(* IEC 61131-3 sources: T4Exjobb/Sigma/Stations/MachineControl/MachineControl/Class/_TCPIP_SERVER (part 2) *)

        (*================================================================*)
        else // - INVALID COMMAND
        (*================================================================*)
          Retcode := TCP_SVR_ERR_SET_PARA_INVALID_CMD;

      end_case;
    else
      Retcode := TCP_SVR_ERR_INVALID_SOCKET;
    end_if;
  else
    Retcode := TCP_SVR_ERR_INVALID_SOCKET;
  end_if;

END_FUNCTION

FUNCTION VIRTUAL GLOBAL _TCPIP_SERVER::ReadMainParameter
	VAR_INPUT
		Cmd 	: DINT;
		SubCmd 	: DINT;
		pParaValue 	: ^DINT;
	END_VAR
	VAR_OUTPUT
		Retcode 	: DINT;
	END_VAR

  Retcode := TCP_SVR_NO_ERROR;

  if (usInit > 0) then
    case Cmd of
      (*================================================================*)
      TCPSVR_CMD_SETSOCKOPT:
      (*================================================================*)
        case SubCmd of
          (*==================================================*)
          TCPSVR_SOCKOPT_NAGLE:
          (*==================================================*)
            if (MainSockOpt.Nagle = false) then
              pParaValue^ := 0;
            else
              pParaValue^ := 1;
            end_if;
          (*==================================================*)
          TCPSVR_SOCKOPT_KEEPALIVE:
          (*==================================================*)
            if (MainSockOpt.KeepAlive = false) then
              pParaValue^ := 0;
            else
              pParaValue^ := 1;
            end_if;
          (*==================================================*)
          TCPSVR_SOCKOPT_DELAYEDACK:
          (*==================================================*)
            if (MainSockOpt.DelayedAck = false) then
              pParaValue^ := 0;
            else
              pParaValue^ := 1;
            end_if;
          (*==================================================*)
          TCPSVR_SOCKOPT_REUSEADDR:
          (*==================================================*)
            if (MainSockOpt.ReuseAddr = false) then
              pParaValue^ := 0;
            else
              pParaValue^ := 1;
            end_if;
          (*==================================================*)
          else // - INVALID SUB COMMAND
          (*==================================================*)
            Retcode := TCP_SVR_ERR_SET_PARA_INVALID_SUB_CMD;
        end_case;

      (*================================================================*)
      TCPSVR_CMD_TASKPRIO:
      (*================================================================*)
        case SubCmd of
          (*==================================================*)
          TCPSVR_SUB_CMD_TASKPRIO:
          (*==================================================*)
            pParaValue^ := AP_TaskPriority$DINT;
          (*==================================================*)
          else // - INVALID SUB COMMAND
          (*==================================================*)
            Retcode := TCP_SVR_ERR_SET_PARA_INVALID_SUB_CMD;
        end_case;

      (*================================================================*)
      TCPSVR_CMD_KEEPALIVEPARA: // - ASYNC TASK PRIORITY
      (*================================================================*)
        case SubCmd of
          (*==================================================*)
          TCPSVR_KEEPALIVE_KEEPIDLE:
          (*==================================================*)
            pParaValue^ := KeepAlivePara.keepIDLE;
          (*==================================================*)
          TCPSVR_KEEPALIVE_KEEPINTVL:
          (*==================================================*)
            pParaValue^ := KeepAlivePara.keepINTVL;
          (*==================================================*)
          TCPSVR_KEEPALIVE_KEEPCNT:
          (*==================================================*)
            pParaValue^ := KeepAlivePara.keepCNT;
          (*==================================================*)
          else // - INVALID SUB COMMAND
          (*==================================================*)
            Retcode := TCP_SVR_ERR_SET_PARA_INVALID_SUB_CMD;
        end_case;

      (*================================================================*)
      TCPSVR_CMD_CLOSESOCKETTYPE:
      (*================================================================*)
        case SubCmd of
          (*==================================================*)
          TCPSVR_CLOSESOCKETTYPE:
          (*==================================================*)
            pParaValue^$UDINT := CloseSocketType;
          (*==================================================*)
          else // - INVALID SUB COMMAND
          (*==================================================*)
            Retcode := TCP_SVR_ERR_SET_PARA_INVALID_SUB_CMD;
        end_case;

      (*================================================================*)
      else // - INVALID COMMAND
      (*================================================================*)
        Retcode := TCP_SVR_ERR_SET_PARA_INVALID_CMD;

    end_case;
  else
    Retcode := TCP_SVR_ERR_MAIN_INIT;
  end_if;

END_FUNCTION

FUNCTION VIRTUAL GLOBAL _TCPIP_SERVER::ReadSocketParameter
	VAR_INPUT
		dSock 	: DINT;
		Cmd 	: DINT;
		SubCmd 	: DINT;
		pParaValue 	: ^DINT;
	END_VAR
	VAR_OUTPUT
		Retcode 	: DINT;
	END_VAR
VAR
	pConn       : ^_CONNECTION;
END_VAR

  Retcode := TCP_SVR_NO_ERROR;

  if (CheckSocketValid(dSock, (#pConn)$^pVoid) = true) then
    if (pConn <> NIL) then
      case Cmd of
        (*================================================================*)
        TCPSVR_CMD_SETSOCKOPT:
        (*================================================================*)
          case SubCmd of
            (*==================================================*)
            TCPSVR_SOCKOPT_NAGLE:
            (*==================================================*)
              if (pConn^.ConnSockOpt.Nagle = false) then
                pParaValue^ := 0;
              else
                pParaValue^ := 1;
              end_if;
            (*==================================================*)
            TCPSVR_SOCKOPT_KEEPALIVE:
            (*==================================================*)
              if (pConn^.ConnSockOpt.KeepAlive = false) then
                pParaValue^ := 0;
              else
                pParaValue^ := 1;
              end_if;
            (*==================================================*)
            TCPSVR_SOCKOPT_DELAYEDACK:
            (*==================================================*)
              if (pConn^.ConnSockOpt.DelayedAck = false) then
                pParaValue^ := 0;
              else
                pParaValue^ := 1;
              end_if;
            (*==================================================*)
            TCPSVR_SOCKOPT_REUSEADDR:
            (*==================================================*)
              if (pConn^.ConnSockOpt.ReuseAddr = false) then
                pParaValue^ := 0;
              else
                pParaValue^ := 1;
              end_if;
            (*==================================================*)
            else // - INVALID SUB COMMAND
            (*==================================================*)
              Retcode := TCP_SVR_ERR_SET_PARA_INVALID_SUB_CMD;
          end_case;

        (*================================================================*)
        TCPSVR_CMD_KEEPALIVEPARA: // - ASYNC TASK PRIORITY
        (*================================================================*)
          case SubCmd of
            (*==================================================*)
            TCPSVR_KEEPALIVE_KEEPIDLE:
            (*==================================================*)
              pParaValue^ := pConn^.KeepAlivePara.keepIDLE;
            (*==================================================*)
            TCPSVR_KEEPALIVE_KEEPINTVL:
            (*==================================================*)
              pParaValue^ := pConn^.KeepAlivePara.keepINTVL;
            (*==================================================*)
            TCPSVR_KEEPALIVE_KEEPCNT:
            (*==================================================*)
              pParaValue^ := pConn^.KeepAlivePara.keepCNT;
            (*==================================================*)
            else // - INVALID SUB COMMAND
            (*==================================================*)
              Retcode := TCP_SVR_ERR_SET_PARA_INVALID_SUB_CMD;
          end_case;

        (*================================================================*)
        TCPSVR_CMD_CLOSESOCKETTYPE:
        (*================================================================*)
          case SubCmd of
            (*==================================================*)
            TCPSVR_CLOSESOCKETTYPE:
            (*==================================================*)
              pParaValue^$UDINT := pConn^.CloseSocketType;
            (*==================================================*)
            else // - INVALID SUB COMMAND
            (*==================================================*)
              Retcode := TCP_SVR_ERR_SET_PARA_INVALID_SUB_CMD;
          end_case;

        (*================================================================*)
        else // - INVALID COMMAND
        (*================================================================*)
          Retcode := TCP_SVR_ERR_SET_PARA_INVALID_CMD;

      end_case;
    else
      Retcode := TCP_SVR_ERR_INVALID_SOCKET;
    end_if;
  else
    Retcode := TCP_SVR_ERR_INVALID_SOCKET;
  end_if;

END_FUNCTION

FUNCTION _TCPIP_SERVER::CheckSocketValid
VAR_INPUT
  dSock 	  : DINT;
  ppConn    : ^pVoid;
END_VAR
VAR_OUTPUT
  Retcode 	: BOOL;
END_VAR
VAR
	i         : USINT;
END_VAR

  Retcode := false;
  if (ppConn <> NIL) then
    ppConn^ := NIL;
  end_if;

  for i := 0 to (MaxConn-1) do
    if (SocketArray[i].dSocket = dSock) then
      if (ppConn <> NIL) then
        ppConn^ := (#SocketArray[i])$^void;
      end_if;
      Retcode := true;
      exit;
    end_if;
  end_for;

END_FUNCTION
